(* PLC project Vn_networks3, Beckhoff Automation GmbH TwinCAT PLC Control 3.5.13.21 *)
(* stored: creationDateTime 1970-01-01T00:00:00 *)

PROGRAM Vn_networks3

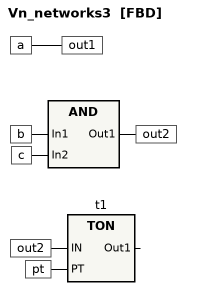
(* FBD diagram, written out as Structured Text *)
out1 := a;
out2 := b AND c;
t1(IN := out2, PT := pt);
END_PROGRAM
